// TIA Portal V21 export
// export: Created 2026-11-07T15:24:57.6561816Z, ExportSetting WithDefaults, DisplayName Totally Integrated Automation Portal, DisplayVersion V21, DisplayName STEP 7 Professional, DisplayVersion V21, DisplayName STEP 7 Safety, DisplayVersion V21, DisplayName Tech WebApplication, DisplayVersion V21, DisplayName WinCC Basic/Comfort/Advanced, DisplayVersion V21, DisplayName WinCC Unified, DisplayVersion V21
Screen "R05_BtnNav"  1024x768, Number=44, Template=Tpl
  ScreenLayer 
    Button "P_NavBtn" at 10,10 size 100x30  Mode=Text, StyleItem=Button, TextOff="BTN", TextOn="BTN"
      on Press: ActivateScreen(Screen name := Alarms, Object number := 0)
